{attribute 'qualified_only'}
{attribute 'strict'}
TYPE E_InterConnection :
(
	NotConnected := 0,
	ConnToTriBlender,
	ConnToLine,
	ConnToTank,
	ConnToCIP
);
END_TYPE

(* stored: Version 1.1.0.1, ProductVersion 3.1.4024.12
   DUT E_InterConnection: Id {9a0727c1-86be-49c5-a623-faa66e7ecd6e} *)
